// Mitsubishi GX Works2 project: 260928   PLC: Q03UDV

PROGRAM MAIN
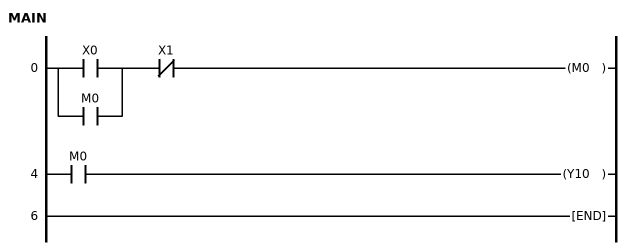
0     LD      X0
      OR      M0
      ANI     X1
      OUT     M0
4     LD      M0
      OUT     Y10
6     END
END_PROGRAM
